Fanuc KAREL source: kx00003.KL

-- PROVISIONAL review KL for V1013-1; original PC SHA256 7af9390c98d3b6f47a705a13f9867c9e3ff8bc529abd2c492864411d4e4e92c8
-- Incomplete behavior may be omitted. Consult companion uncertainty JSON. Do not deploy.
PROGRAM KX00003
%NOLOCKGROUP
VAR
  I : INTEGER
  J : INTEGER
  B : BOOLEAN
  F : FILE
  S : STRING[80]
-- UNRESOLVED_DECL P type=000102
BEGIN
  -- UNRESOLVED_PC offsets 5-32; opcodes 22,3F,3F,3D
  -- UNRESOLVED_PC offsets 37-65; opcodes 22,3F,9C,9C,37,9C,9C,37,2C
  -- UNRESOLVED_PC offsets 70-77; opcodes 22,39
  -- UNRESOLVED_PC offsets 82-86; opcodes 7F
END KX00003
